// TIA Portal V20 export
// export: Created 2026-10-20T18:54:11.7686072Z, ExportSetting None, DisplayName Totally Integrated Automation Portal, DisplayVersion V20 Update 6, DisplayName TIA Portal Openness, DisplayVersion V20 Update 6, DisplayName TIA Portal Version Control Interface, DisplayVersion V20 Update 6, DisplayName SINAMICS Startdrive Advanced, DisplayVersion V20 SP1, DisplayName SINAMICS Startdrive G130, G150, S120, S150, SINAMICS MV, G220, S200, S210, DisplayVersion V20 SP1, DisplayName SINAMICS Startdrive G110M, G120, G120C, G120D, G120P, G115D, DisplayVersion V20 SP1, DisplayName STEP 7 Professional, DisplayVersion V20 Update 6, DisplayName STEP 7 Safety, DisplayVersion V20 Update 2, DisplayName WinCC Basic/Comfort/Advanced, DisplayVersion V20 Update 6, DisplayName WinCC Unified, DisplayVersion V20 Update 6
VAR_GLOBAL   // PLC tag table "Errors"
   "Sick Lector_Error code 2" AT %MW748 : Word;
   Errors_Profinet_2 AT %MW732 : Word;
   "IND_360_SB Status Group 1" AT %MW742 : Word;
   Errors_IND360_Smart5_Red_Level_5 AT %MW700 : Word;
   Errors_Profinet_1 AT %MW730 : Word;
   "Sick Lector_Error code 1" AT %MW746 : Word;
   Error AT %M729.0 : Bool;
   Errors_Profinet_3 AT %MW734 : Word;
   Errors_Profinet_4 AT %MW754 : Word;
   Errors_Profinet_5 AT %MW756 : Word;
   Errors_Profinet_9 AT %MW764 : Word;
   Errors_Profinet_8 AT %MW762 : Word;
   Errors_Profinet_7 AT %MW760 : Word;
   Erros_Supply_Feedback_5 AT %MW768 : Word;
   Erros_Supply_Feedback_7 AT %MW772 : Word;
   Erros_Supply_Feedback_6 AT %MW770 : Word;
   Erros_Supply_Feedback_4 AT %MW766 : Word;
   Errors_Profinet_6 AT %MW758 : Word;
   Erros_Supply_Feedback_1 AT %MW736 : Word;
   Erros_Supply_Feedback_2 AT %MW738 : Word;
   Erros_Supply_Feedback_3 AT %MW740 : Word;
   "Sick Lector_Error code 3" AT %MW790 : Word;
   "Sick Lector_Error code 5" AT %MW794 : Word;
   "Sick Lector_Error code 4_2" AT %MW802 : Word;
   "Linear Encoder_Device Errors 4" AT %MW778 : Word;
   "Linear Encoder_Warnings 5" AT %MW788 : Word;
   "Linear Encoder_Device Errors 3" AT %MW776 : Word;
   "Linear Encoder_Warnings 3" AT %MW784 : Word;
   "Sick Lector_Error code 4" AT %MW792 : Word;
   "Sick Lector_Error code 2_2" AT %MW798 : Word;
   "Linear Encoder_Device Errors 2" AT %MW774 : Word;
   "Linear Encoder_Warnings 2" AT %MW782 : Word;
   "Linear Encoder_Device Errors 5" AT %MW780 : Word;
   "Sick Lector_Error code 1_2" AT %MW796 : Word;
   "Sick Lector_Error code 3_2" AT %MW800 : Word;
   "Sick Lector_Error code 5_2" AT %MW804 : Word;
   "Linear Encoder_Warnings 4" AT %MW786 : Word;
   "Linear Encoder_Device Errors 1" AT %MW750 : Word;
   "Linear Encoder_Warnings 1" AT %MW752 : Word;
   Estop_Error_Word_1 AT %MW808 : Word;
   Estop_Error_Word_3 AT %MW812 : Word;
   Estop_Error_Word_2 AT %MW810 : Word;
   Errors_Profinet_10 AT %MW806 : Word;
   Estop_Error_Word_4 AT %MW814 : Word;
   Estop_Error_Word_5 AT %MW816 : Word;
   Errors_Word_Shuttles_1 AT %MW818 : Word;
   Errors_Word_Shuttles_2 AT %MW820 : Word;
   Errors_Word_Gates_1 AT %MW822 : Word;
   Estop_Error_Word_6 AT %MW824 : Word;
   Errors_Profinet_11 AT %MW826 : Word;
   Errors_Word_LightGuard_1 AT %MW828 : Word;
   Errors_Word_Logistex AT %MW830 : Word;
   Erros_Word_OPC_5 AT %MW840 : Word;
   Erros_Word_OPC_3 AT %MW836 : Word;
   Erros_Word_OPC_4 AT %MW838 : Word;
   Erros_Word_OPC_2 AT %MW834 : Word;
   Erros_Word_OPC_1 AT %MW832 : Word;
   Errors_Word_Gates_2 AT %MW842 : Word;
   Error_MQTT_2 AT %MW846 : Word;
   Error_MQTT AT %MW844 : Word;
   Error_Word_Overhang AT %MW848 : Word;
END_VAR
